TYPE ET_MC_RampType :
(
	ET_MC_RampType_eMTTrapez,
	ET_MC_RampType_eMTSinSquare,
	ET_MC_RampType_eMTParabolic
	
);
END_TYPE

(* stored: Version 1.1.0.1, ProductVersion 3.1.4024.15
   DUT ET_MC_RampType: Id {a20ef4c2-b14f-4504-b029-3dd014478ff7} *)
